Fanuc KAREL source: KT00785.KL

PROGRAM KT00785
%NOLOCKGROUP
VAR
  I1: INTEGER
  I2: INTEGER
  OUT: REAL
BEGIN
  I1 = 2
  I2 = 3
  I1 = 2
  I2 = 3
  OUT = COS(I1)
END KT00785
